// TIA Portal V20 export
// export: Created 2026-10-19T18:45:39.4268706Z, ExportSetting None, DisplayName Totally Integrated Automation Portal, DisplayVersion V20 Update 6, DisplayName TIA Portal Openness, DisplayVersion V20 Update 6, DisplayName TIA Portal Version Control Interface, DisplayVersion V20 Update 6, DisplayName SINAMICS Startdrive Advanced, DisplayVersion V20 SP1, DisplayName SINAMICS Startdrive G130, G150, S120, S150, SINAMICS MV, G220, S200, S210, DisplayVersion V20 SP1, DisplayName SINAMICS Startdrive G110M, G120, G120C, G120D, G120P, G115D, DisplayVersion V20 SP1, DisplayName STEP 7 Professional, DisplayVersion V20 Update 6, DisplayName STEP 7 Safety, DisplayVersion V20 Update 2, DisplayName WinCC Basic/Comfort/Advanced, DisplayVersion V20 Update 6, DisplayName WinCC Unified, DisplayVersion V20 Update 6
VAR_GLOBAL   // PLC tag table "IO_ET200_2"
   "VTD2 LEVEL DETECT 2" AT %I202.1 : Bool;
   "OVERTRAVEL UPPER LIMIT - CH1(2)" AT %I1476.1 : Bool;
   "VTD2 DOCKING PINS 2 EXTEND" AT %Q181.5 : Bool;
   "C2103 STOPPER RAISED" AT %I95.0 : Bool;
   "VTD2 DOCKING PINS EXTENDED 2" AT %I141.1 : Bool;
   "VTD2 DOCKING PINS RETRACTED 2" AT %I141.2 : Bool;
   "C2104 STOPPER LOWERED" AT %I132.1 : Bool;
   "C2102 STOPPER RAISED" AT %I94.0 : Bool;
   "C2103 STOPPER MOTOR" AT %Q95.4 : Bool;
   "VTD2 DOCKING PINS 1 RETRACT" AT %Q181.6 : Bool;
   "OVERTRAVEL LOWER LIMIT - CH2(2)" AT %I1476.4 : Bool;
   "C2105 STOPPER MOTOR" AT %Q133.4 : Bool;
   "C2105 STOPPER LOWERED" AT %I133.1 : Bool;
   "VTD2 DOCKING PINS 1 EXTEND" AT %Q181.4 : Bool;
   "C2104 STOPPER RAISED" AT %I132.0 : Bool;
   "C2105 STOPPER RAISED" AT %I133.0 : Bool;
   "OVERTRAVEL LOWER LIMIT - CH1(2)" AT %I1476.0 : Bool;
   "C2106 STOPPER LOWERED" AT %I140.1 : Bool;
   "VTD2 LEVEL DETECT 1" AT %I202.0 : Bool;
   "C2106 STOPPER RAISED" AT %I140.0 : Bool;
   "VTD2 DOCKING PINS EXTENDED 1" AT %I141.0 : Bool;
   "C2104 STOPPER MOTOR" AT %Q132.4 : Bool;
   "C2102 STOPPER LOWERED" AT %I94.1 : Bool;
   "OVERTRAVEL UPPER LIMIT - CH2(2)" AT %I1476.5 : Bool;
   "C2103 STOPPER LOWERED" AT %I95.1 : Bool;
   "C2106 STOPPER MOTOR" AT %Q140.4 : Bool;
   "VTD2 DOCKING PINS 2 RETRACT" AT %Q181.7 : Bool;
   "C2102 STOPPER MOTOR" AT %Q94.4 : Bool;
   "VTD2 DOCKING PINS RETRACTED 1" AT %I141.3 : Bool;
END_VAR
